FUNCTION_BLOCK MODE_SM
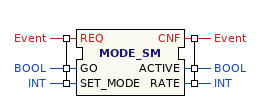
  EVENT_INPUT
    REQ WITH GO, SET_MODE;
  END_EVENT
  EVENT_OUTPUT
    CNF WITH ACTIVE, RATE;
  END_EVENT
  VAR_INPUT
    GO : BOOL;
    SET_MODE : INT;
  END_VAR
  VAR_OUTPUT
    ACTIVE : BOOL;
    RATE : INT;
  END_VAR
  VAR
    GAIN : INT;
  END_VAR
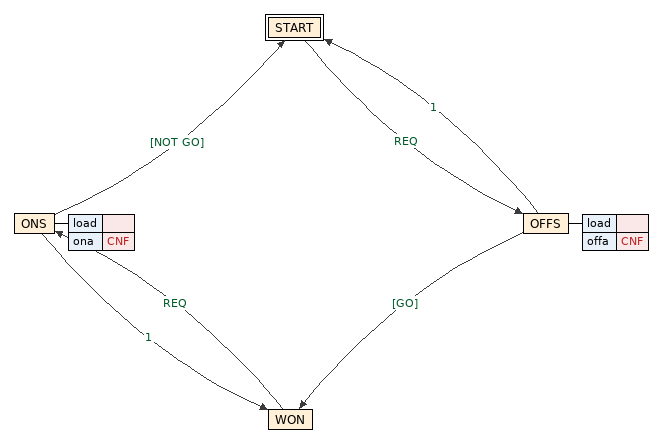
  EC_STATES
    START;
    OFFS : load, offa -> CNF;
    WON;
    ONS : load, ona -> CNF;
  END_STATES
  EC_TRANSITIONS
    START TO OFFS := REQ;
    OFFS TO WON := [GO];
    OFFS TO START := 1;
    WON TO ONS := REQ;
    ONS TO START := [NOT GO];
    ONS TO WON := 1;
  END_TRANSITIONS
  ALGORITHM load IN ST:
IF SET_MODE <> 0 THEN GAIN := SET_MODE; END_IF;
  END_ALGORITHM
  ALGORITHM offa IN ST:
CASE GAIN OF 1: RATE := 0; 2: RATE := 100; END_CASE;
IF GO THEN ACTIVE := TRUE; END_IF;
  END_ALGORITHM
  ALGORITHM ona IN ST:
CASE GAIN OF 1: RATE := RATE + 1; 2: RATE := RATE + 2; END_CASE;
IF NOT GO THEN ACTIVE := FALSE; END_IF;
  END_ALGORITHM
END_FUNCTION_BLOCK
